Fanuc KAREL source: kt00891.KL

PROGRAM KT00891
%STACKSIZE=65535
%PRIORITY=65535
%NOLOCKGROUP
VAR
P1 : JOINTPOS9
P2 : JOINTPOS9
OUT : POSITION
BEGIN
-- UNRESOLVED_PC line 8 opcodes [27 27 49 7E AD 76 7E 4A] marker_code=0
END KT00891
